(* CODESYS project counter.library
   DefaultNamespace: KOSTAL.AF2024.Misc.Counter
   DocFormat: reStructuredText
   Description: Component to handle/store counter data in several formats
   Author: M. Hundt / Frank Dümpelmann
   Title: KOSTAL.AF2024.Misc.Counter
   Version: 1.0.1.0
   Company: KOSTAL GmbH & Co.KG
   Placeholder: KOSTAL.AF2024.Misc.Counter

Project tree, tasks and I/O mapping:
  libraries: KOSTAL.AF2024.Core.ID, 1.0.0.0 (KOSTAL GmbH & Co.KG); KOSTAL.AF2024.Core.JsonTools, 1.0.0.0 (KOSTAL GmbH & Co.KG); KOSTAL.AF2024.Core.Process, 1.0.0.0 (KOSTAL GmbH & Co.KG); KOSTAL.AF2024.Core.Settings, 1.0.0.0 (KOSTAL GmbH & Co.KG); KOSTAL.AF2024.Core.Station, 1.0.0.0 (KOSTAL GmbH & Co.KG); KOSTAL.AF2024.Core.StringTools, 1.0.0.0 (KOSTAL GmbH & Co.KG); KOSTAL.AF2024.Core.System, 1.0.0.0 (KOSTAL GmbH & Co.KG); KOSTAL.AF2024.HMI.I_Hmi, 1.0.0.0 (KOSTAL GmbH & Co.KG); Tc2_Standard, 3.3.3.0 (Beckhoff Automation GmbH); Tc2_System, 3.6.2.0 (Beckhoff Automation GmbH)
  0_Counter/
    function block _FB_Counter [ST]: Counter, INC, Init, Reset, toString
    interface _I_Counter: Counter, INC, Init, Reset, toString
    interface _I_Counter_RO: Counter, toString
  1_CounterSet/
    interface I_T_CounterSet: Fail, Pass
    function block T_CounterSet [ST]: Fail, Pass
  2_Base/
    function block _FB_Base [ST]: _HMI_define, _parameterControl, _resetCondition, _storage, LinkStorage, Fail, Pass, ResetEnable, FBmain
    data type E_text_counter
  3_Storage/
    0_Interface/
      DUT/
        interface I_StorageContent: Clear, CopyFrom, CopyTo, Fail, Pass
        interface I_StorageContent_CopyFrom: CopyFrom
        interface I_StorageContent_RO: CopyTo, Fail, Pass
        function block T_StorageContent [ST]: Clear, CopyFrom, CopyTo, Fail, Pass
      interface I_Storage: Content, Reset, State
    1_Json/
      function block FB_Json [ST]: _Step_ClearContent, _Step_CreateContent, _Step_Finish, _Step_Idle_EXT, _Step_ParseContent, _hasContentChanged, Content, Reset, State, storageMode, FBmain
  Project Information/
    function F_GetCompany [ST]
    function F_GetTitle [ST]
    function F_GetVersion [ST]
  Version/
    global variables Global_Version
  data type E_FileMode
  data type E_StorageMode
*)

// 2_Base/E_text_counter
{attribute 'qualified_only'}
{attribute 'strict'}
TYPE E_text_counter :
(
	Language:= 1,
	myName	:= 2,
	PASS		:= 3,
	FAIL		:= 4,
	
	manualReset			:= 10,
	automaticReset	:= 11,
	
	RESET	:= 100
);
END_TYPE

// E_FileMode
{attribute 'qualified_only'}
{attribute 'strict'}
TYPE E_FileMode :
(
	Idle := 0,
	ReadFile,
	WriteFile
);
END_TYPE

// E_StorageMode
{attribute 'qualified_only'}
{attribute 'strict'}
TYPE E_StorageMode :
(
	file := 0,
	web
);
END_TYPE

// Version/Global_Version
{attribute 'TcGenerated'}
{attribute 'no-analysis'}
{attribute 'linkalways'}
// This function has been automatically generated from the project information.
VAR_GLOBAL CONSTANT
	{attribute 'const_non_replaced'}
	stLibVersion_KOSTAL_AF2024_Misc_Counter : ST_LibVersion := (iMajor := 1, iMinor := 0, iBuild := 1, iRevision := 0, nFlags := 0, sVersion := '1.0.1.0');
END_VAR

// 0_Counter/_FB_Counter
FUNCTION_BLOCK _FB_Counter IMPLEMENTS _I_Counter, _I_Counter_RO
VAR
	_Counter	: UDINT;	//UDINT
END_VAR

PROPERTY PUBLIC Counter : UDINT
GET

Counter:= _Counter;
END_GET
END_PROPERTY

METHOD PUBLIC INC : BOOL

IF _counter + 1 < _counter THEN	RETURN;	END_IF

_Counter:= _Counter + 1;

INC:= TRUE;
END_METHOD

METHOD PUBLIC Init
VAR_INPUT
	value	: UDINT;	// UDINT
END_VAR

_Counter:= value;
END_METHOD

METHOD PUBLIC Reset
VAR_INPUT
END_VAR

_Counter:= UDINT#0;
END_METHOD

METHOD PUBLIC toString : STRING

toString:= UDINT_TO_STRING(_Counter);
END_METHOD

END_FUNCTION_BLOCK

// 0_Counter/_I_Counter
INTERFACE _I_Counter EXTENDS KOSTAL_AF2024_Core_System.I_Interface

PROPERTY PUBLIC Counter : UDINT
GET
END_GET
END_PROPERTY

METHOD PUBLIC INC : BOOL
END_METHOD

METHOD PUBLIC Init
VAR_INPUT
	value	: UDINT;	// UDINT
END_VAR
END_METHOD

METHOD PUBLIC Reset
VAR_INPUT
END_VAR
END_METHOD

METHOD PUBLIC toString : STRING
END_METHOD

END_INTERFACE

// 0_Counter/_I_Counter_RO
INTERFACE _I_Counter_RO EXTENDS KOSTAL_AF2024_Core_System.I_Interface

PROPERTY PUBLIC Counter : UDINT
GET
END_GET
END_PROPERTY

METHOD PUBLIC toString : STRING
VAR_INPUT
END_VAR
END_METHOD

END_INTERFACE

// 1_CounterSet/I_T_CounterSet
INTERFACE I_T_CounterSet

PROPERTY Fail : _I_Counter
GET
END_GET
END_PROPERTY

PROPERTY Pass : _I_Counter
GET
END_GET
END_PROPERTY

END_INTERFACE

// 1_CounterSet/T_CounterSet
FUNCTION_BLOCK PUBLIC T_CounterSet IMPLEMENTS I_T_CounterSet
VAR
	_Pass	:	_FB_Counter;
	_Fail	:	_FB_Counter;
END_VAR

PROPERTY Fail : _I_Counter
GET

Fail:= _Fail;
END_GET
END_PROPERTY

PROPERTY Pass : _I_Counter
GET

Pass:= _Pass;
END_GET
END_PROPERTY

END_FUNCTION_BLOCK

// 2_Base/_FB_Base
(* 
:Author: Martin Hundt <m.hundt@kostal.com>,  
:Date: 2021-11-11
 
Function 
======== 
| Base class for a good part/bad part counter
| Reads Data from I_CounterStorage interface
| Provides I_Counter interface to the application
 
 
Methods and Properties
===========================
| Icounter_Pass/Icounter_Fail: Access to the counters - Increase, reset and read value
| link_IcounterStorage: Link a storage component with the I_Storage interface
| ResetEnable: Disable reset of the counter (e.g. set true in manual mode)
| FBmain(): To be called cyclically 

 
Usage sample: 
============= 
| See best practice
 
*)

FUNCTION_BLOCK ABSTRACT _FB_Base EXTENDS KOSTAL_AF2024_Core_Station.FB_Station_Free IMPLEMENTS I_T_CounterSet

VAR

	//=======================================================================================================================================
	//_ID	: KOSTAL_AF2024_Core_ID.FB_ID;

	
	//===========================================================================================================
	//Interfaces
	//===========================================================================================================

//	_condition	: KOSTAL_AF2024_Core_Process.FB_processCondition;
//	_state			: KOSTAL_AF2024_Core_Process.FB_plcState;
	
	//_languageAvailable	: BOOL;
	
	//HMI
	_pageStation		: KOSTAL_AF2024_HMI_I_Hmi.I_Page_Station_Owner; 

	_resetEnable		: BOOL;
	//_message			: KOSTAL_AF2024_Core_Process.FB_messageText_3_lines;
	
	//===========================================================================================================
	//I_Counter
	_counterPass	: _FB_Counter;
	_counterFail	: _FB_Counter;

	//===========================================================================================================
	//I_CounterStorage
	_Istorage							: I_Storage;
	_initFromStorageDone	: BOOL:= FALSE;	// BOOL


END_VAR

METHOD PROTECTED _HMI_define
VAR_INPUT
END_VAR

_pageStation.Name:= "Counter";

_pageStation.Text.line_01:= _condition.message.line_01;
_pageStation.Text.line_02:= _condition.message.line_02;
_pageStation.Text.line_03:= _condition.message.line_03;
 
_pageStation.Button_Escape.Visible	:= _condition.isError();
_pageStation.Button_Escape.Text		:= "Reset";
          
_pageStation.Button_OnOff.Visible	:= _resetEnable;
_pageStation.Button_OnOff.Text			:= "RESET";
          
_pageStation.Status.CopyFrom(_condition);
          
//default 
_pageStation.Buttons_Custom.Button(1).Visible	:= FALSE;
_pageStation.Buttons_Custom.Button(2).Visible	:= FALSE;
END_METHOD

METHOD Protected _parameterControl : BOOL
VAR_INPUT
END_VAR

_parameterControl:= FALSE;

IF _Istorage = 0 THEN

	_message.clear();
	_message.line_01:= "Parameter Fail";
	_message.line_02:= "Interface _I_storage is not linked";

	_condition.setMessage(4999, _message);

ELSE
	
	_parameterControl:= TRUE;

END_IF
END_METHOD

METHOD PROTECTED _resetCondition
VAR_INPUT
END_VAR

IF _condition.isInfo() THEN
	_condition.clear();
ELSIF _condition.isText() THEN
	_condition.clear();
ELSIF _condition.isMessage() THEN
	_condition.clear();
ELSIF _condition.isMasterMessage() THEN
	_condition.clear();
ELSIF _pageStation.Button_Escape.Pulse THEN
	_condition.clear();
END_IF
END_METHOD

METHOD PROTECTED _storage
VAR_INPUT
END_VAR


IF	_Istorage.State.fail THEN

	_message.clear();
	_message.line_01:= "ERROR Counter Storage";
	_message.line_02:= _Istorage.State.description;

	_condition.setMessage(_condition.PriorityLevel_Error, _message);
	
	IF _pageStation.Button_Escape.Pulse THEN
		 _Istorage.Reset();
	END_IF

ELSIF NOT _Istorage.State.ready THEN

	_message.clear();
	_message.line_01:= "wait for Counter Storage >Ready<";
	_message.line_02:= _Istorage.State.description;
	
	_condition.setMessage(_condition.PriorityLevel_Message, _message);


ELSIF NOT _initFromStorageDone THEN

	_counterPass.Init(_Istorage.Content.Pass);
	_counterFail.Init(_Istorage.Content.Fail);
	
	_initFromStorageDone:= TRUE;
	
ELSE	
	_Istorage.Content.fail:= _counterFail.Counter;
	_Istorage.Content.Pass:= _counterPass.Counter;
	
	_message.clear();
	_message.line_01:= "Counter is ready";
	_message.line_02:= _Istorage.State.description;
	_condition.setMessage(_condition.PriorityLevel_Info, _message);
END_IF
END_METHOD

METHOD PUBLIC LinkStorage
VAR_INPUT
	link	: I_Storage;
END_VAR

_Istorage:= link;
END_METHOD

PROPERTY Fail : _I_Counter
GET

Fail:= _counterFail;
END_GET
END_PROPERTY

PROPERTY Pass : _I_Counter
GET

Pass:= _counterPass;
END_GET
END_PROPERTY

//Set true to enable reset button on HMI
PROPERTY ResetEnable : BOOL
GET
ResetEnable := _resetEnable;
END_GET
SET
_resetEnable := ResetEnable;
END_SET
END_PROPERTY

METHOD PUBLIC FBmain
VAR_INPUT
END_VAR

IF NOT _parameterControl() THEN RETURN;	END_IF

_HMI_define();

_resetCondition();

_storage();
END_METHOD

END_FUNCTION_BLOCK

// 3_Storage/0_Interface/I_Storage
INTERFACE I_Storage EXTENDS KOSTAL_AF2024_Core_System.I_Interface

PROPERTY Content : I_StorageContent
GET
END_GET
END_PROPERTY

METHOD Reset	: BOOL
END_METHOD

PROPERTY State : KOSTAL_AF2024_Core_Process.I_T_plcState
GET
END_GET
END_PROPERTY

END_INTERFACE

// 3_Storage/0_Interface/DUT/I_StorageContent
INTERFACE I_StorageContent EXTENDS KOSTAL_AF2024_Core_System.I_Interface

METHOD PUBLIC Clear
END_METHOD

METHOD PUBLIC CopyFrom
VAR_INPUT
	IN	: I_StorageContent_RO;
END_VAR
END_METHOD

METHOD PUBLIC CopyTo
VAR_INPUT
	IN	: I_StorageContent_CopyFrom;
END_VAR
END_METHOD

PROPERTY PUBLIC Fail : UDINT
GET
END_GET
SET
END_SET
END_PROPERTY

PROPERTY PUBLIC Pass : UDINT
GET
END_GET
SET
END_SET
END_PROPERTY

END_INTERFACE

// 3_Storage/0_Interface/DUT/I_StorageContent_RO
INTERFACE I_StorageContent_RO EXTENDS KOSTAL_AF2024_Core_System.I_Interface

METHOD PUBLIC CopyTo
VAR_INPUT
	IN	: I_StorageContent_CopyFrom;
END_VAR
END_METHOD

PROPERTY PUBLIC Fail : UDINT
GET
END_GET
END_PROPERTY

PROPERTY PUBLIC Pass : UDINT
GET
END_GET
END_PROPERTY

END_INTERFACE

// 3_Storage/0_Interface/DUT/I_StorageContent_CopyFrom
INTERFACE I_StorageContent_CopyFrom EXTENDS KOSTAL_AF2024_Core_System.I_Interface

METHOD PUBLIC CopyFrom
VAR_INPUT
	IN	: I_StorageContent_RO;
END_VAR
END_METHOD

END_INTERFACE

// 3_Storage/0_Interface/DUT/T_StorageContent
FUNCTION_BLOCK T_StorageContent IMPLEMENTS I_StorageContent, I_StorageContent_RO, I_StorageContent_CopyFrom
VAR
	_Pass	: UDINT;
	_Fail	: UDINT;
END_VAR

METHOD PUBLIC Clear

_Pass:= UDINT#0;
_Fail:= UDINT#0;
END_METHOD

METHOD PUBLIC CopyFrom
VAR_INPUT
	IN	: I_StorageContent_RO;
END_VAR

IF IN = 0 THEN RETURN;	END_IF

_Pass:= IN.Pass;
_Fail:= IN.Fail;
END_METHOD

METHOD PUBLIC CopyTo
VAR_INPUT
	IN	: I_StorageContent_CopyFrom;
END_VAR

IF IN = 0 THEN RETURN;	END_IF

IN.CopyFrom(THIS^);
END_METHOD

PROPERTY PUBLIC Fail : UDINT
GET

Fail:= _Fail;
END_GET
SET

_Fail:= Fail;
END_SET
END_PROPERTY

PROPERTY PUBLIC Pass : UDINT
GET

Pass:= _Pass;
END_GET
SET

_Pass:= Pass;
END_SET
END_PROPERTY

END_FUNCTION_BLOCK

// 3_Storage/1_Json/FB_Json
(* 
:Author: Martin Hundt <m.hundt@kostal.com>,  
:Date: 2021-11-11
 
Function 
======== 
| Stores counter values in a json file and provides it to a counter component via the ICounterStorage interface
| The file is loaded when the application starts and is stored when a counter value changed
 
 
Methods and Properties
===========================
| fullQualifiedFile: Path to the storage file
| FBmain(): To be called cyclically
| IcounterStorage_Content(.pass/.fail): value of the counters (Part of I_CounterStorage interface)
| IcounterStorage_Status: Status of the component: ready = file loaded correctly, fail = file loading failed  
 

 
Usage sample: 
============= 
| Also see counter best practice
 
.. code::  
 
 PROGRAM MAIN 
 VAR 
 	_counter		: Kostal_TC3_Components_Counter_FlexHMI.FB_Counter;
	_counterStorage : Kostal_TC3_Components_Counter_Storage_Json.FB_Storage;
 END_VAR 
  
 	//Define Counter Storage
	_counterStorage.fullQualifiedFile := 'C:\test\counter.json';
	_counterStorage.FBmain();
	
	//Define Counter and link Counter Storage
	_counter.link_IcounterStorage(_counterStorage);
	_counter.FBmain();
 
*)

FUNCTION_BLOCK PUBLIC FB_Json EXTENDS KOSTAL_AF2024_Core_JsonTools._FB_Base IMPLEMENTS I_Storage
VAR

	_mode							: E_FileMode;
	_content					: T_StorageContent;	
	_contentAsLoaded	: T_StorageContent;
	_reset						: BOOL;
	_init							: BOOL:= TRUE;

	
	//file handling
	//_stepJson		: KOSTAL_AF2024_Core_Process.FB_processStep_Flow;	
	
	
	//storage mode
	_storageMode	: E_StorageMode:= E_StorageMode.file;	//default file mode is set

END_VAR

VAR CONSTANT
	_MEMBERNAME_PASS 	: STRING := 'PASSPARTS';
	_MEMBERNAME_FAIL	: STRING := 'FAILPARTS';

	_COUNTER_ADDRESS_ERROR	: INT:= 10;
END_VAR

(*
	Overwrite to clear your data content before parse content
*)
METHOD PROTECTED _Step_ClearContent


_content.Clear();
_contentAsLoaded.Clear();

SUPER^._Step_ClearContent();
END_METHOD

(*
	Overwrite to create your data content
*)
METHOD PROTECTED _Step_CreateContent

VAR
	_string: STRING;
END_VAR

_NewDocument();

_string:= UDINT_TO_STRING(_content.Pass);
_parser.AddStringMember(_jDoc, _MEMBERNAME_PASS, _string);

_string:= UDINT_TO_STRING(_content.Fail);
_parser.AddStringMember(_jDoc, _MEMBERNAME_FAIL, _string);

SUPER^._Step_CreateContent();
END_METHOD

METHOD PROTECTED _Step_Finish : BOOL
VAR_INPUT
END_VAR


SUPER^._Step_Finish();

_contentAsLoaded.CopyFrom(_content);

_Step.set(0);
END_METHOD

(*
	Overwrite to add your Idle content here
*)
METHOD PROTECTED _Step_Idle_EXT : BOOL
VAR_INPUT
END_VAR

_Step_Idle_EXT:= FALSE;

IF _storageMode = E_StorageMode.file AND _fullQualifiedFile = '' THEN

	_Step_Idle_EXT:= TRUE;

	_State.clear();
	_State.fail:= TRUE;
	_State.description:= "ERROR - no filename defined";

ELSIF _storageMode = E_StorageMode.web AND 	_extFileName = '' THEN

	_Step_Idle_EXT:= TRUE;

	_State.clear();
	_State.fail:= TRUE;
	_State.description:= "ERROR - no extended filename defined";
	
ELSIF _storageMode = E_StorageMode.web AND 	_extFilePath = '' THEN

	_Step_Idle_EXT:= TRUE;

	_State.clear();
	_State.fail:= TRUE;
	_State.description:= "ERROR - no extended filepath defined";

ELSIF _DocumentIsEmpty() THEN

	IF _storageMode = E_StorageMode.file	THEN	_THIS_CALLED:= E_THIS_CALLED.FILE_READ;
	ELSE																				_THIS_CALLED:= E_THIS_CALLED.WEB_READ;
	END_IF

ELSIF _hasContentChanged() THEN

	IF _storageMode = E_StorageMode.file	THEN	_THIS_CALLED:= E_THIS_CALLED.FILE_WRITE;
	ELSE																				_THIS_CALLED:= E_THIS_CALLED.WEB_WRITE;
	END_IF

ELSE	_THIS_CALLED:= E_THIS_CALLED.IDL;

END_IF
END_METHOD

(*
	Overwrite to parse your data content
*)
METHOD PROTECTED _Step_ParseContent

_content.pass := _PARSE_UDINT(_jDoc,_MEMBERNAME_PASS, FALSE, 0);
_content.Fail := _PARSE_UDINT(_jDoc,_MEMBERNAME_FAIL, FALSE, 0);


SUPER^._Step_ParseContent();
END_METHOD

METHOD PROTECTED _hasContentChanged : BOOL

_hasContentChanged:=		(_content.Pass <> _contentAsLoaded.Pass)
										OR	(_content.Fail <> _contentAsLoaded.Fail);



//(Tc2_System.MEMCMP(ADR(_CompCompare), ADR(_CompContent), SIZEOF(_CompContent)) <> 0);
END_METHOD

PROPERTY Content : I_StorageContent
GET

Content:= _content;
END_GET
END_PROPERTY

METHOD Reset	: BOOL

_Step.init();
END_METHOD

PROPERTY State : KOSTAL_AF2024_Core_Process.I_T_plcState
GET

State:= SUPER^._State;
END_GET
END_PROPERTY

PROPERTY PUBLIC storageMode : E_StorageMode
GET

storageMode:= _storageMode;
END_GET
SET

_storageMode:= storageMode;
END_SET
END_PROPERTY

METHOD PUBLIC FBmain

//_a0_Setting();

//_stepJson.Header();

//IF _stepJson.isActive(0)	THEN	_a10_Origin();	END_IF
//IF _stepJson.isActive(1)	THEN	_a20_ReadContent();		END_IF

//IF _stepJson.NotFound()		THEN	_a1_Fail();			END_IF


//IF _content = 0 THEN
//	_State.clear();
//	_State.fail:= TRUE;
//	_State.description:= "no Counter content is linked";
//	RETURN;
//END_IF

//IF _DocumentIsEmpty() THEN
	
//END_IF

SUPER^._FBmain();
 
_init:= FALSE;
END_METHOD

END_FUNCTION_BLOCK

// Project Information/F_GetCompany
// This function has been automatically generated from the project information.
{attribute 'signature_flag' := '1073741824'}
{attribute 'TcGenerated'}
{attribute 'no-analysis'}
FUNCTION F_GetCompany : WSTRING
VAR_INPUT
	
END_VAR

F_GetCompany := "KOSTAL GmbH & Co.KG";

END_FUNCTION

// Project Information/F_GetTitle
// This function has been automatically generated from the project information.
{attribute 'signature_flag' := '1073741824'}
{attribute 'TcGenerated'}
{attribute 'no-analysis'}
FUNCTION F_GetTitle : WSTRING
VAR_INPUT
	
END_VAR

F_GetTitle := "KOSTAL.AF2024.Misc.Counter";

END_FUNCTION

// Project Information/F_GetVersion
// This function has been automatically generated from the project information.
{attribute 'signature_flag' := '1073741824'}
{attribute 'TcGenerated'}
{attribute 'no-analysis'}
FUNCTION F_GetVersion : ST_LibVersion
VAR_INPUT
	
END_VAR

F_GetVersion.iMajor := 1;
F_GetVersion.iMinor := 0;
F_GetVersion.iBuild := 1;
F_GetVersion.iRevision := 0;
F_GetVersion.sVersion := '1.0.1.0';
F_GetVersion.nFlags := 0;

END_FUNCTION
